FUNCTION_BLOCK FB_VFD_Drive_REF
VAR_INPUT
	stTerminalState			AT %I*:ST_TerminalState;
	stVfdToPlc				AT %I*:ST_VFDTOPLC;
	stPlcToVfd				AT %Q*:ST_PLCTOVFD;
END_VAR
VAR_OUTPUT

END_VAR
VAR_IN_OUT

END_VAR
VAR

END_VAR

;

END_FUNCTION_BLOCK

(* stored: Version 1.1.0.1, ProductVersion 3.1.4024.15
   POU FB_VFD_Drive_REF: Id {7f68e1f5-fe9d-481a-9640-a8628c98594c}, SpecialFunc None *)
